Fanuc KAREL source: kb00178.compact.KL

PROGRAM KB00178
%STACKSIZE=65535
%PRIORITY=65535
%NOLOCKGROUP
%ENVIRONMENT REGOPE
VAR
P1 : INTEGER
P2 : REAL
P3 : INTEGER
BEGIN
P1=1
P2=1.0
P3=1
SET_REAL_REG(P1,P2,P3)
END KB00178
